(* Logix 5000 project; controller CIP_14485201 vendor 1 type 14 code 216 rev 38.11; software revision 38.01; part 9 of 12 *)
(* tags used below, declared in another part *)
   Bit : BOOL[128];   // BIT
   MOA_OFF : DINT[20];   // PANELVIEW MOA OFF
   MOA_ON : DINT[20];   // PANELVIEW MOA ON
   OpCode_Pin : DINT[5];   // OPCODE PIN ARRAY
   Panelview : INT[40];   // PANELVIEW CONTROL
   PID2 : PID;   // SUPPLY FLOW PID
   PID2_bumpless_transfer : BOOL;   // FORCE PID TO RESTART FROM PREVIOUS OUTPUT VALUE
   PID2_Man_Mode : BOOL;   // PID2 MANUAL MODE
   PID2_Manual_PB_Pressed : BOOL;   // PID2 MANUAL PUSHBUTTON PRESSED
   PID2_Output_Memory : REAL;   // SUPPLY FLOW PID OUTPUT MEMORY TO USE FOR BUMPLESS TRANSFER
   PID2_PV_Manual_PB : BOOL;   // PID2 MANUAL MODE SELECTED ON HMI
   PID2_Setpoint_Memory : REAL;   // SUPPLY FLOW PID SETPOINT MEMORY TO USE FOR BUMPLESS TRANSFER
   PID_Ons : DINT[6];   // PID ONE SHOT
   PID_Timer : TIMER[5];   // PID TIMERS
   PV_Output_Status : INT[20];   // PV OUTPUT STATUS:
   PV_Output_Status_IND : INT[20,16];   // PV OUTPUT STATUS IND:
   PV_Status_Bit : BOOL;   // SYSTEM BIT
   Recipe : RECIPE[41];   // RECIPES
   SP_Supply_Flow : REAL;   // CURRENT SUPPLY FLOW SETPOINT
   Supply_Mod_Valve_force_open : BOOL;   // FORCE SUPPLY MOD. VALVE TO 100% OPEN
   Utility_Button : DINT[5];   // PANELVIEW UTILITY BUTTONS
   Utility_Button_Ons : DINT[5];   // PANELVIEW UTILITY BUTTON ONE SHOTS
   Utility_Ons : DINT[5];   // PANELVIEW UTILITY ONE SHOTS
   Utility_Out : DINT[5];   // PANELVIEW UTILITY OUTPUT CONTROL
   Utility_Timer : TIMER[4];   // PANELVIEW UTILITY TIMERS
(* MainProgram, continued *)

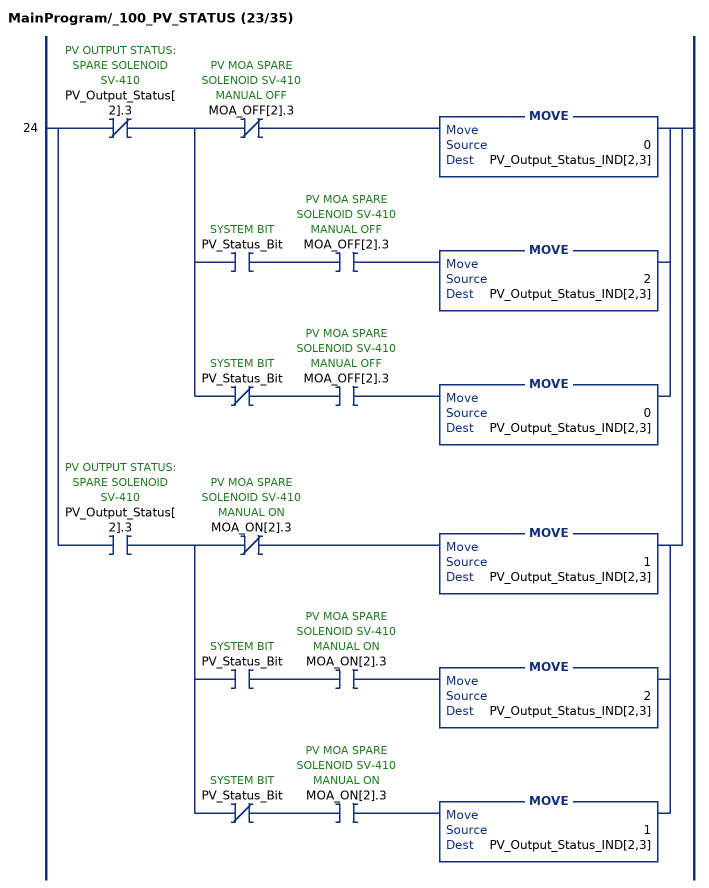
   [picture p140: MainProgram/_100_PV_STATUS rungs 24-24]
   24: [XIO(PV_Output_Status[2].3) [XIO(MOA_OFF[2].3) MOVE(0,PV_Output_Status_IND[2,3]) ,XIC(PV_Status_Bit) XIC(MOA_OFF[2].3) MOVE(2,PV_Output_Status_IND[2,3]) ,XIO(PV_Status_Bit) XIC(MOA_OFF[2].3) MOVE(0,PV_Output_Status_IND[2,3]) ] ,XIC(PV_Output_Status[2].3) [XIO(MOA_ON[2].3) MOVE(1,PV_Output_Status_IND[2,3]) ,XIC(PV_Status_Bit) XIC(MOA_ON[2].3) MOVE(2,PV_Output_Status_IND[2,3]) ,XIO(PV_Status_Bit) XIC(MOA_ON[2].3) MOVE(1,PV_Output_Status_IND[2,3]) ] ];
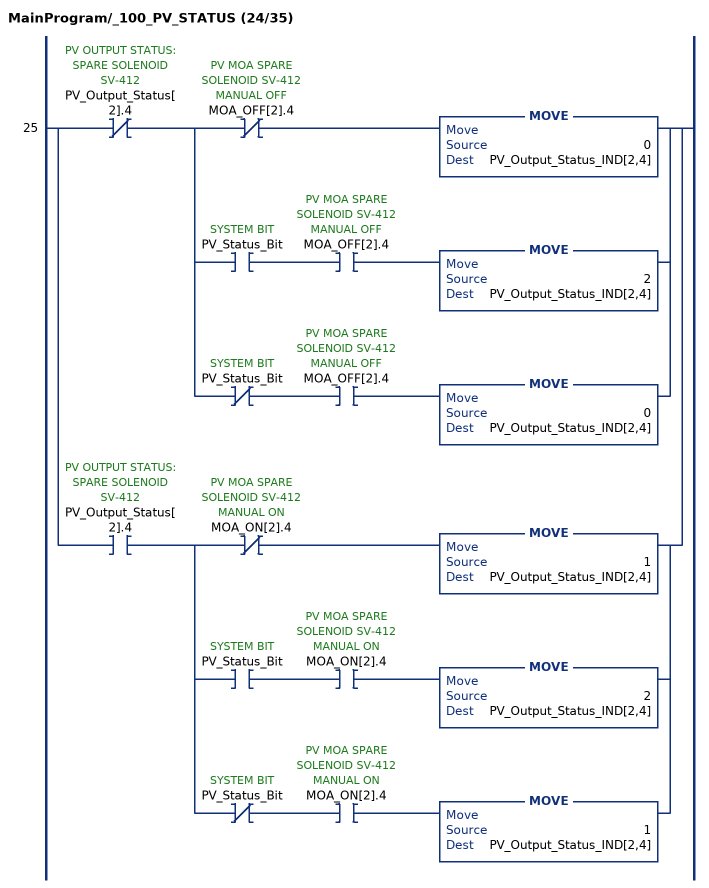
   25: [XIO(PV_Output_Status[2].4) [XIO(MOA_OFF[2].4) MOVE(0,PV_Output_Status_IND[2,4]) ,XIC(PV_Status_Bit) XIC(MOA_OFF[2].4) MOVE(2,PV_Output_Status_IND[2,4]) ,XIO(PV_Status_Bit) XIC(MOA_OFF[2].4) MOVE(0,PV_Output_Status_IND[2,4]) ] ,XIC(PV_Output_Status[2].4) [XIO(MOA_ON[2].4) MOVE(1,PV_Output_Status_IND[2,4]) ,XIC(PV_Status_Bit) XIC(MOA_ON[2].4) MOVE(2,PV_Output_Status_IND[2,4]) ,XIO(PV_Status_Bit) XIC(MOA_ON[2].4) MOVE(1,PV_Output_Status_IND[2,4]) ] ];
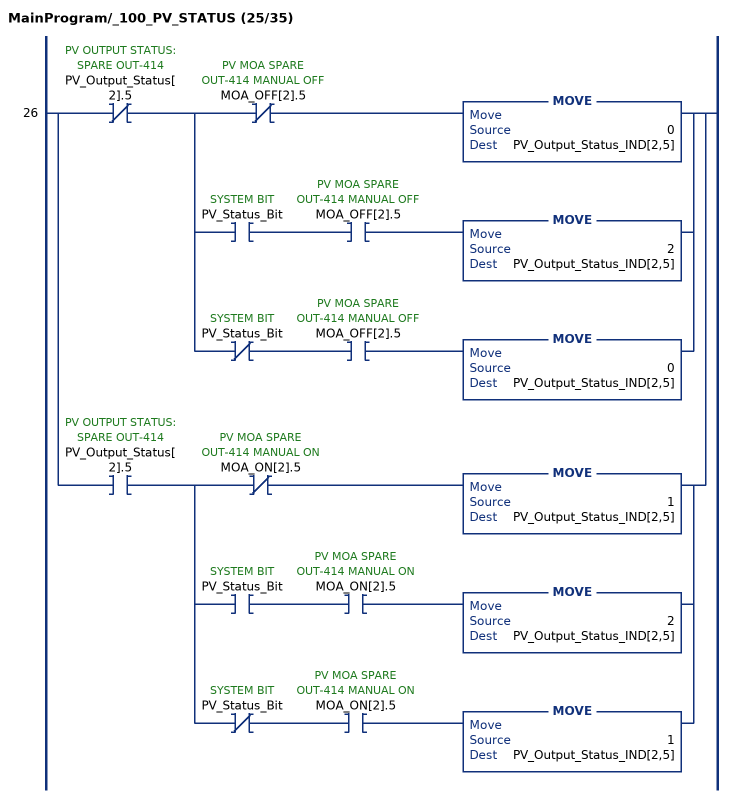
   26: [XIO(PV_Output_Status[2].5) [XIO(MOA_OFF[2].5) MOVE(0,PV_Output_Status_IND[2,5]) ,XIC(PV_Status_Bit) XIC(MOA_OFF[2].5) MOVE(2,PV_Output_Status_IND[2,5]) ,XIO(PV_Status_Bit) XIC(MOA_OFF[2].5) MOVE(0,PV_Output_Status_IND[2,5]) ] ,XIC(PV_Output_Status[2].5) [XIO(MOA_ON[2].5) MOVE(1,PV_Output_Status_IND[2,5]) ,XIC(PV_Status_Bit) XIC(MOA_ON[2].5) MOVE(2,PV_Output_Status_IND[2,5]) ,XIO(PV_Status_Bit) XIC(MOA_ON[2].5) MOVE(1,PV_Output_Status_IND[2,5]) ] ];
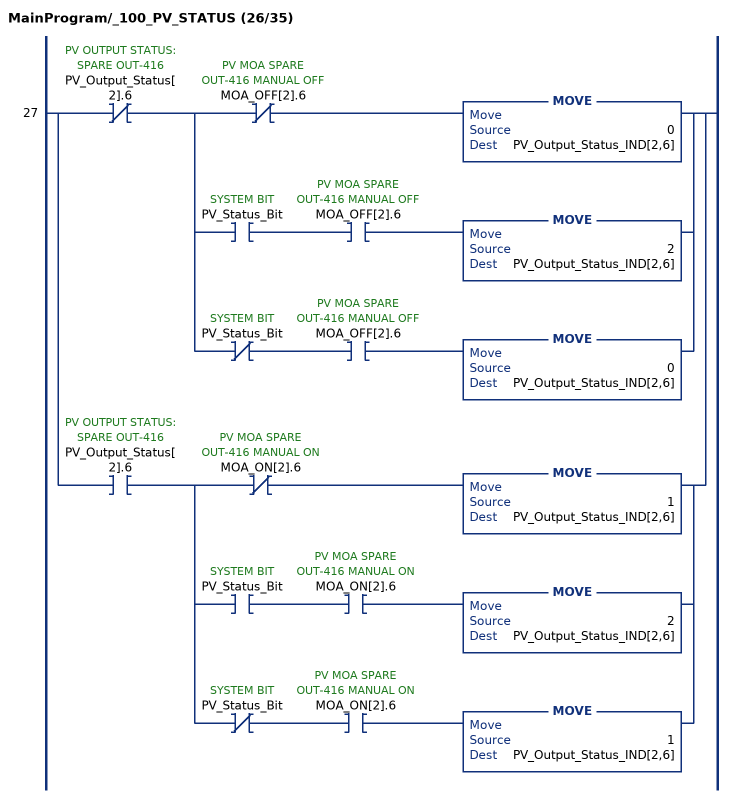
   27: [XIO(PV_Output_Status[2].6) [XIO(MOA_OFF[2].6) MOVE(0,PV_Output_Status_IND[2,6]) ,XIC(PV_Status_Bit) XIC(MOA_OFF[2].6) MOVE(2,PV_Output_Status_IND[2,6]) ,XIO(PV_Status_Bit) XIC(MOA_OFF[2].6) MOVE(0,PV_Output_Status_IND[2,6]) ] ,XIC(PV_Output_Status[2].6) [XIO(MOA_ON[2].6) MOVE(1,PV_Output_Status_IND[2,6]) ,XIC(PV_Status_Bit) XIC(MOA_ON[2].6) MOVE(2,PV_Output_Status_IND[2,6]) ,XIO(PV_Status_Bit) XIC(MOA_ON[2].6) MOVE(1,PV_Output_Status_IND[2,6]) ] ];
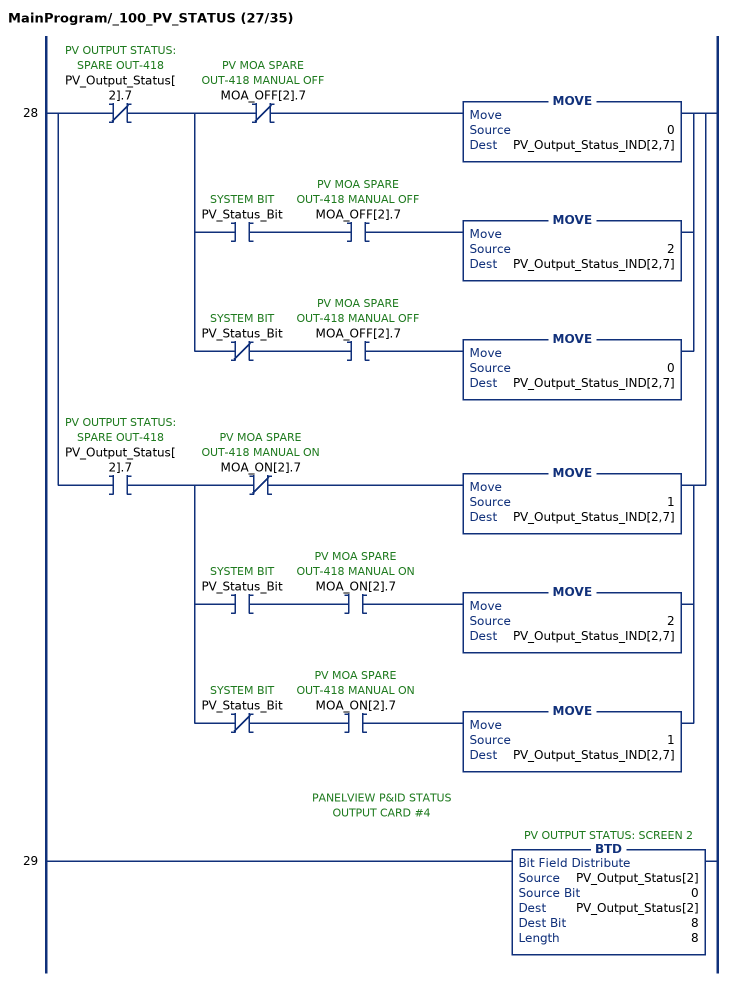
   28: [XIO(PV_Output_Status[2].7) [XIO(MOA_OFF[2].7) MOVE(0,PV_Output_Status_IND[2,7]) ,XIC(PV_Status_Bit) XIC(MOA_OFF[2].7) MOVE(2,PV_Output_Status_IND[2,7]) ,XIO(PV_Status_Bit) XIC(MOA_OFF[2].7) MOVE(0,PV_Output_Status_IND[2,7]) ] ,XIC(PV_Output_Status[2].7) [XIO(MOA_ON[2].7) MOVE(1,PV_Output_Status_IND[2,7]) ,XIC(PV_Status_Bit) XIC(MOA_ON[2].7) MOVE(2,PV_Output_Status_IND[2,7]) ,XIO(PV_Status_Bit) XIC(MOA_ON[2].7) MOVE(1,PV_Output_Status_IND[2,7]) ] ];
   // PANELVIEW P&ID STATUS
   // OUTPUT CARD #4
   29: BTD(PV_Output_Status[2],0,PV_Output_Status[2],8,8);
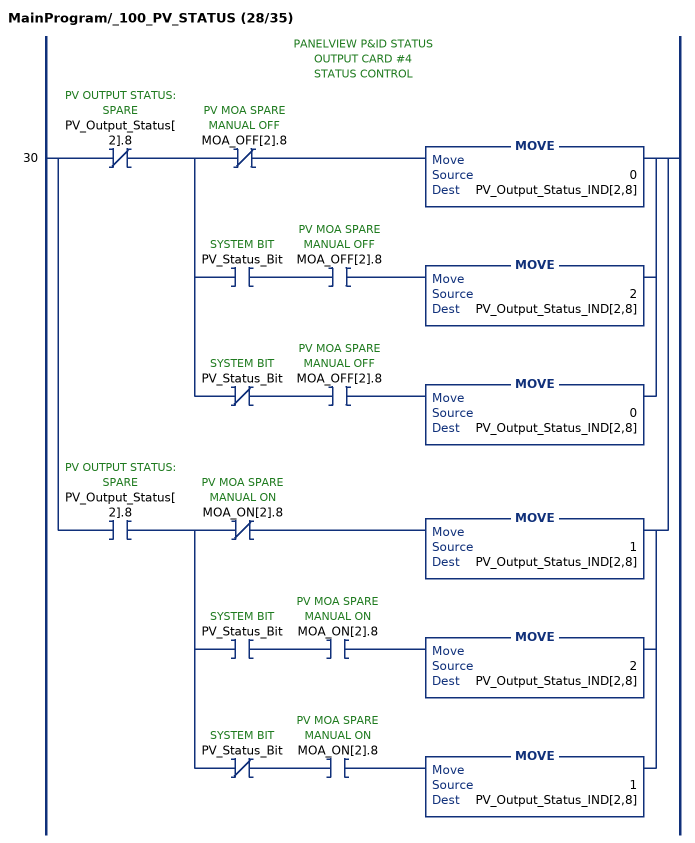
   // PANELVIEW P&ID STATUS
   // OUTPUT CARD #4
   // STATUS CONTROL
   30: [XIO(PV_Output_Status[2].8) [XIO(MOA_OFF[2].8) MOVE(0,PV_Output_Status_IND[2,8]) ,XIC(PV_Status_Bit) XIC(MOA_OFF[2].8) MOVE(2,PV_Output_Status_IND[2,8]) ,XIO(PV_Status_Bit) XIC(MOA_OFF[2].8) MOVE(0,PV_Output_Status_IND[2,8]) ] ,XIC(PV_Output_Status[2].8) [XIO(MOA_ON[2].8) MOVE(1,PV_Output_Status_IND[2,8]) ,XIC(PV_Status_Bit) XIC(MOA_ON[2].8) MOVE(2,PV_Output_Status_IND[2,8]) ,XIO(PV_Status_Bit) XIC(MOA_ON[2].8) MOVE(1,PV_Output_Status_IND[2,8]) ] ];
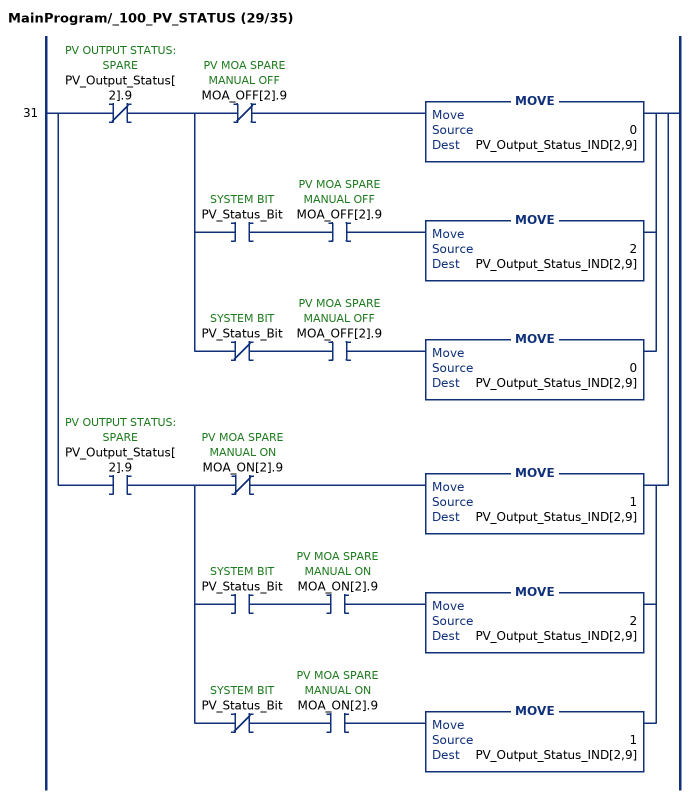
   31: [XIO(PV_Output_Status[2].9) [XIO(MOA_OFF[2].9) MOVE(0,PV_Output_Status_IND[2,9]) ,XIC(PV_Status_Bit) XIC(MOA_OFF[2].9) MOVE(2,PV_Output_Status_IND[2,9]) ,XIO(PV_Status_Bit) XIC(MOA_OFF[2].9) MOVE(0,PV_Output_Status_IND[2,9]) ] ,XIC(PV_Output_Status[2].9) [XIO(MOA_ON[2].9) MOVE(1,PV_Output_Status_IND[2,9]) ,XIC(PV_Status_Bit) XIC(MOA_ON[2].9) MOVE(2,PV_Output_Status_IND[2,9]) ,XIO(PV_Status_Bit) XIC(MOA_ON[2].9) MOVE(1,PV_Output_Status_IND[2,9]) ] ];
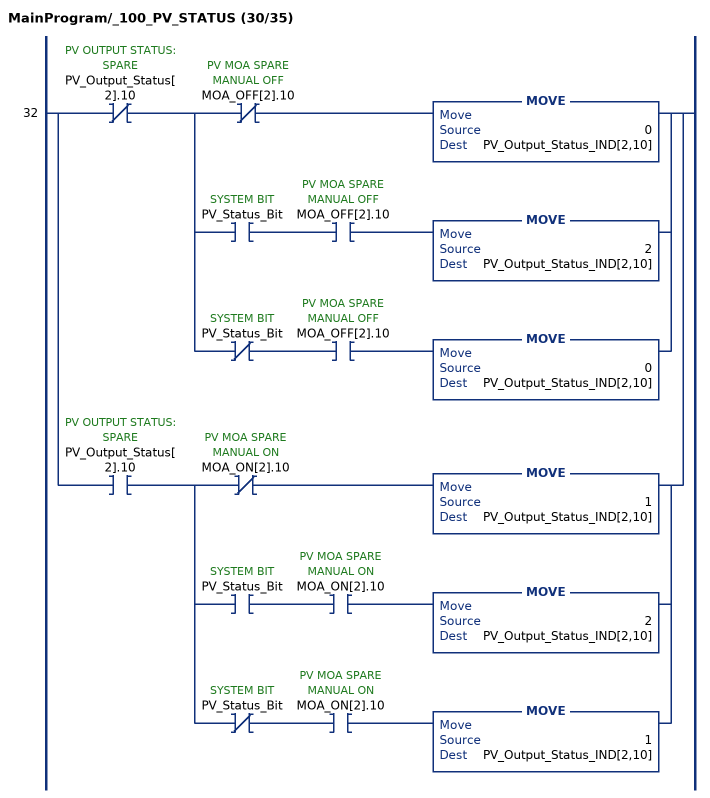
   32: [XIO(PV_Output_Status[2].10) [XIO(MOA_OFF[2].10) MOVE(0,PV_Output_Status_IND[2,10]) ,XIC(PV_Status_Bit) XIC(MOA_OFF[2].10) MOVE(2,PV_Output_Status_IND[2,10]) ,XIO(PV_Status_Bit) XIC(MOA_OFF[2].10) MOVE(0,PV_Output_Status_IND[2,10]) ] ,XIC(PV_Output_Status[2].10) [XIO(MOA_ON[2].10) MOVE(1,PV_Output_Status_IND[2,10]) ,XIC(PV_Status_Bit) XIC(MOA_ON[2].10) MOVE(2,PV_Output_Status_IND[2,10]) ,XIO(PV_Status_Bit) XIC(MOA_ON[2].10) MOVE(1,PV_Output_Status_IND[2,10]) ] ];
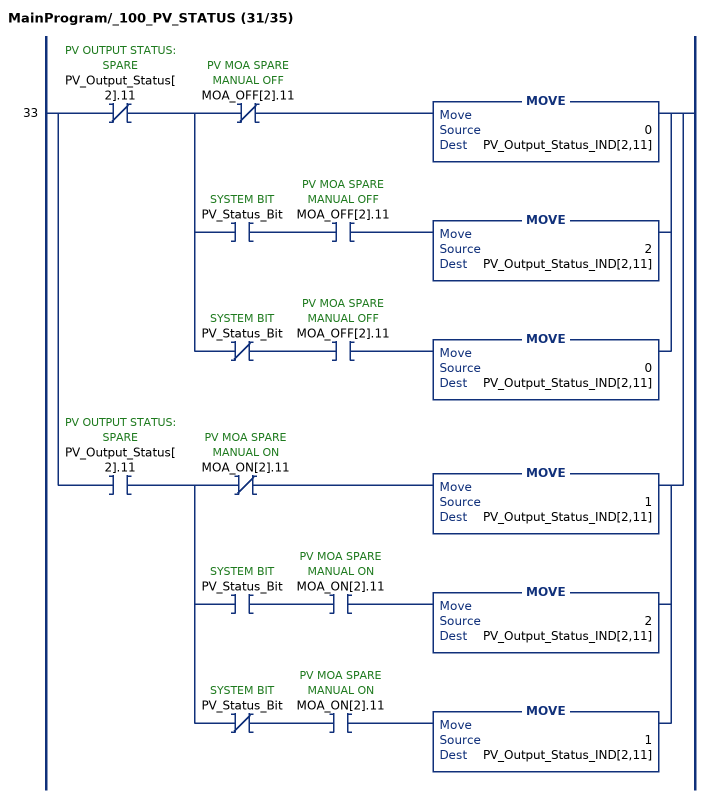
   33: [XIO(PV_Output_Status[2].11) [XIO(MOA_OFF[2].11) MOVE(0,PV_Output_Status_IND[2,11]) ,XIC(PV_Status_Bit) XIC(MOA_OFF[2].11) MOVE(2,PV_Output_Status_IND[2,11]) ,XIO(PV_Status_Bit) XIC(MOA_OFF[2].11) MOVE(0,PV_Output_Status_IND[2,11]) ] ,XIC(PV_Output_Status[2].11) [XIO(MOA_ON[2].11) MOVE(1,PV_Output_Status_IND[2,11]) ,XIC(PV_Status_Bit) XIC(MOA_ON[2].11) MOVE(2,PV_Output_Status_IND[2,11]) ,XIO(PV_Status_Bit) XIC(MOA_ON[2].11) MOVE(1,PV_Output_Status_IND[2,11]) ] ];
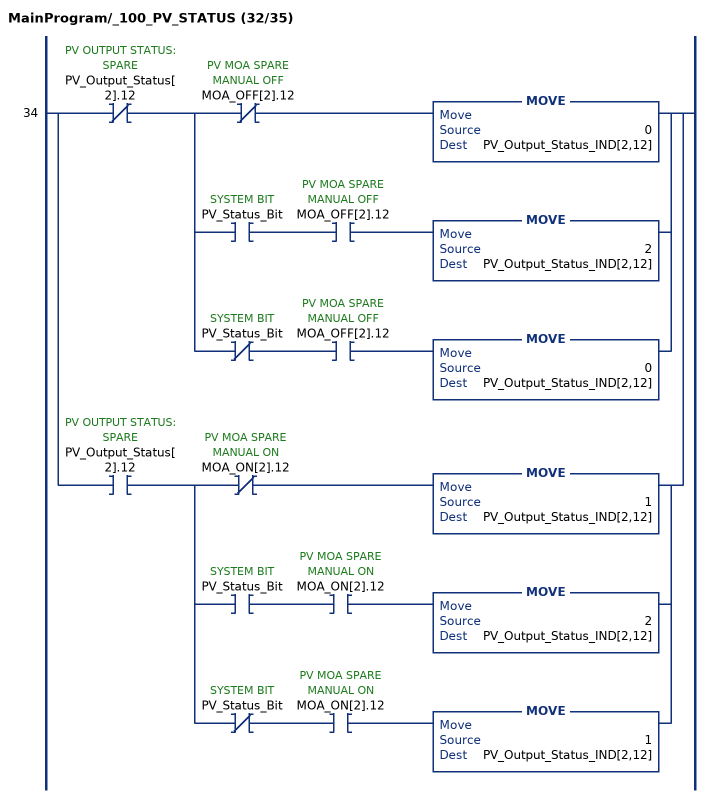
   34: [XIO(PV_Output_Status[2].12) [XIO(MOA_OFF[2].12) MOVE(0,PV_Output_Status_IND[2,12]) ,XIC(PV_Status_Bit) XIC(MOA_OFF[2].12) MOVE(2,PV_Output_Status_IND[2,12]) ,XIO(PV_Status_Bit) XIC(MOA_OFF[2].12) MOVE(0,PV_Output_Status_IND[2,12]) ] ,XIC(PV_Output_Status[2].12) [XIO(MOA_ON[2].12) MOVE(1,PV_Output_Status_IND[2,12]) ,XIC(PV_Status_Bit) XIC(MOA_ON[2].12) MOVE(2,PV_Output_Status_IND[2,12]) ,XIO(PV_Status_Bit) XIC(MOA_ON[2].12) MOVE(1,PV_Output_Status_IND[2,12]) ] ];
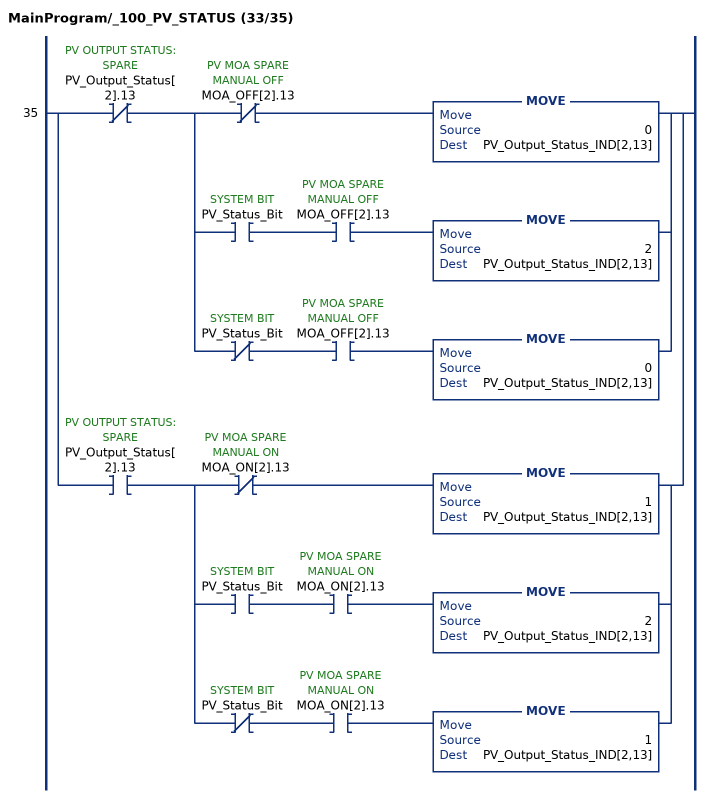
   35: [XIO(PV_Output_Status[2].13) [XIO(MOA_OFF[2].13) MOVE(0,PV_Output_Status_IND[2,13]) ,XIC(PV_Status_Bit) XIC(MOA_OFF[2].13) MOVE(2,PV_Output_Status_IND[2,13]) ,XIO(PV_Status_Bit) XIC(MOA_OFF[2].13) MOVE(0,PV_Output_Status_IND[2,13]) ] ,XIC(PV_Output_Status[2].13) [XIO(MOA_ON[2].13) MOVE(1,PV_Output_Status_IND[2,13]) ,XIC(PV_Status_Bit) XIC(MOA_ON[2].13) MOVE(2,PV_Output_Status_IND[2,13]) ,XIO(PV_Status_Bit) XIC(MOA_ON[2].13) MOVE(1,PV_Output_Status_IND[2,13]) ] ];
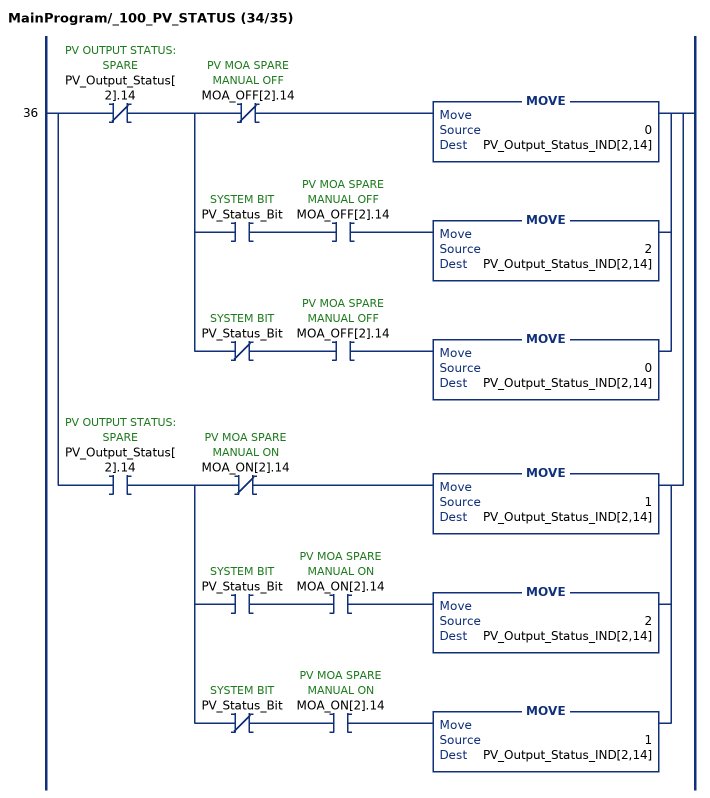
   36: [XIO(PV_Output_Status[2].14) [XIO(MOA_OFF[2].14) MOVE(0,PV_Output_Status_IND[2,14]) ,XIC(PV_Status_Bit) XIC(MOA_OFF[2].14) MOVE(2,PV_Output_Status_IND[2,14]) ,XIO(PV_Status_Bit) XIC(MOA_OFF[2].14) MOVE(0,PV_Output_Status_IND[2,14]) ] ,XIC(PV_Output_Status[2].14) [XIO(MOA_ON[2].14) MOVE(1,PV_Output_Status_IND[2,14]) ,XIC(PV_Status_Bit) XIC(MOA_ON[2].14) MOVE(2,PV_Output_Status_IND[2,14]) ,XIO(PV_Status_Bit) XIC(MOA_ON[2].14) MOVE(1,PV_Output_Status_IND[2,14]) ] ];
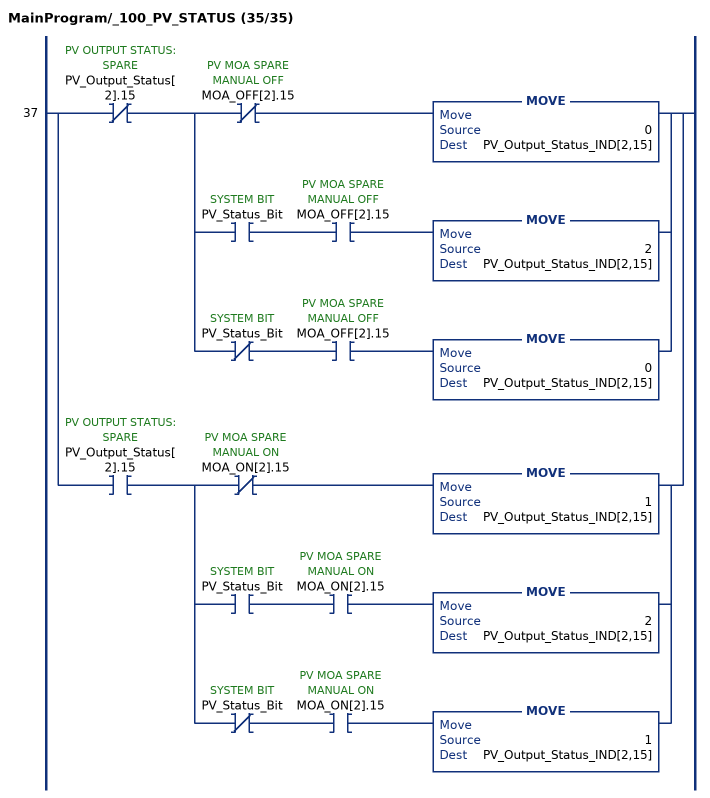
   37: [XIO(PV_Output_Status[2].15) [XIO(MOA_OFF[2].15) MOVE(0,PV_Output_Status_IND[2,15]) ,XIC(PV_Status_Bit) XIC(MOA_OFF[2].15) MOVE(2,PV_Output_Status_IND[2,15]) ,XIO(PV_Status_Bit) XIC(MOA_OFF[2].15) MOVE(0,PV_Output_Status_IND[2,15]) ] ,XIC(PV_Output_Status[2].15) [XIO(MOA_ON[2].15) MOVE(1,PV_Output_Status_IND[2,15]) ,XIC(PV_Status_Bit) XIC(MOA_ON[2].15) MOVE(2,PV_Output_Status_IND[2,15]) ,XIO(PV_Status_Bit) XIC(MOA_ON[2].15) MOVE(1,PV_Output_Status_IND[2,15]) ] ];
END_ROUTINE

ROUTINE _20_UTILITY   (* ladder *)
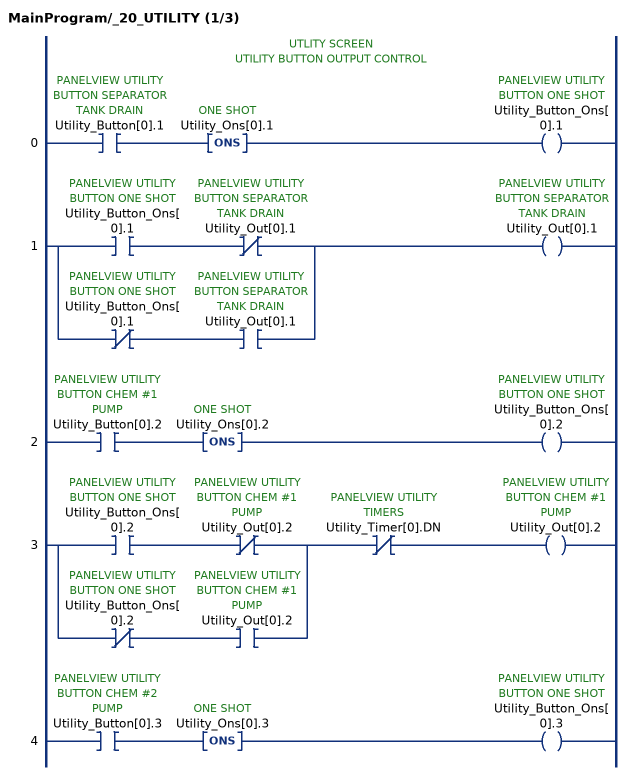
   // UTLITY SCREEN
   // UTILITY BUTTON OUTPUT CONTROL
   0: XIC(Utility_Button[0].1)ONS(Utility_Ons[0].1)OTE(Utility_Button_Ons[0].1);
   1: [XIC(Utility_Button_Ons[0].1) XIO(Utility_Out[0].1) ,XIO(Utility_Button_Ons[0].1) XIC(Utility_Out[0].1) ]OTE(Utility_Out[0].1);
   2: XIC(Utility_Button[0].2)ONS(Utility_Ons[0].2)OTE(Utility_Button_Ons[0].2);
   3: [XIC(Utility_Button_Ons[0].2) XIO(Utility_Out[0].2) ,XIO(Utility_Button_Ons[0].2) XIC(Utility_Out[0].2) ]XIO(Utility_Timer[0].DN)OTE(Utility_Out[0].2);
   4: XIC(Utility_Button[0].3)ONS(Utility_Ons[0].3)OTE(Utility_Button_Ons[0].3);
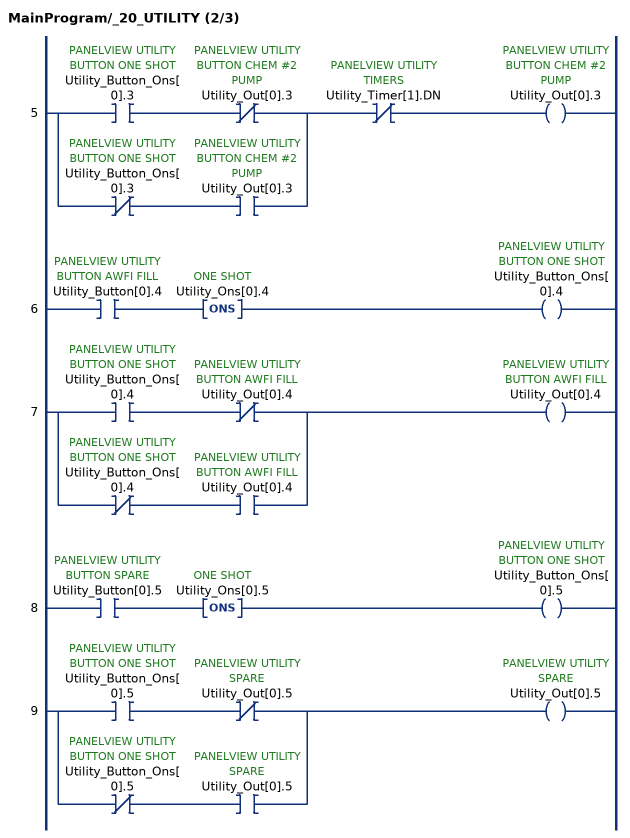
   5: [XIC(Utility_Button_Ons[0].3) XIO(Utility_Out[0].3) ,XIO(Utility_Button_Ons[0].3) XIC(Utility_Out[0].3) ]XIO(Utility_Timer[1].DN)OTE(Utility_Out[0].3);
   6: XIC(Utility_Button[0].4)ONS(Utility_Ons[0].4)OTE(Utility_Button_Ons[0].4);
   7: [XIC(Utility_Button_Ons[0].4) XIO(Utility_Out[0].4) ,XIO(Utility_Button_Ons[0].4) XIC(Utility_Out[0].4) ]OTE(Utility_Out[0].4);
   8: XIC(Utility_Button[0].5)ONS(Utility_Ons[0].5)OTE(Utility_Button_Ons[0].5);
   9: [XIC(Utility_Button_Ons[0].5) XIO(Utility_Out[0].5) ,XIO(Utility_Button_Ons[0].5) XIC(Utility_Out[0].5) ]OTE(Utility_Out[0].5);
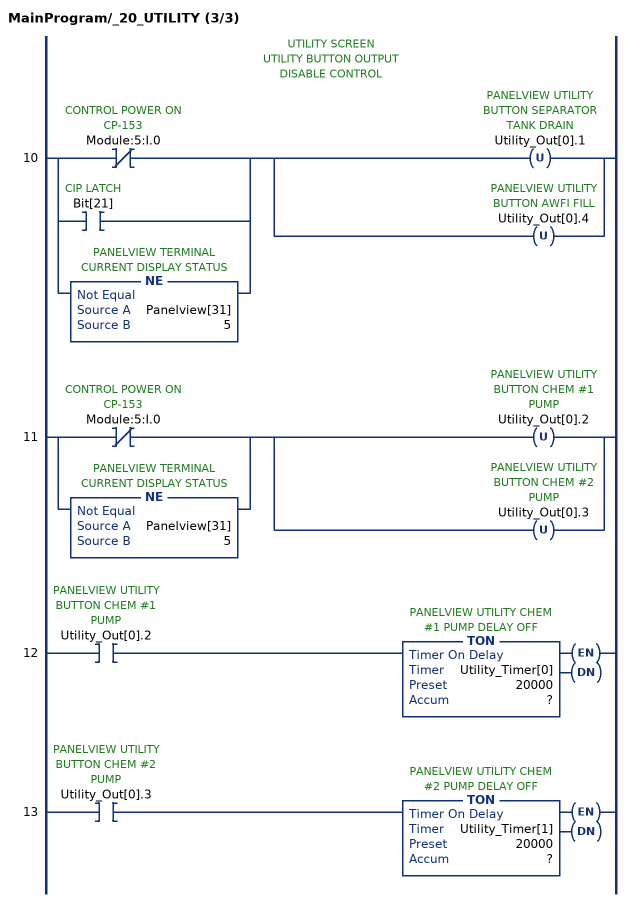
   // UTILITY SCREEN
   // UTILITY BUTTON OUTPUT
   // DISABLE CONTROL
   10: [XIO(Module:5:I.0) ,XIC(Bit[21]) ,NE(Panelview[31],5) ][OTU(Utility_Out[0].1) ,OTU(Utility_Out[0].4) ];
   11: [XIO(Module:5:I.0) ,NE(Panelview[31],5) ][OTU(Utility_Out[0].2) ,OTU(Utility_Out[0].3) ];
   12: XIC(Utility_Out[0].2)TON(Utility_Timer[0],?,?);
   13: XIC(Utility_Out[0].3)TON(Utility_Timer[1],?,?);
END_ROUTINE

ROUTINE _25_PID_SUPPLY_FLOW   (* ladder *)
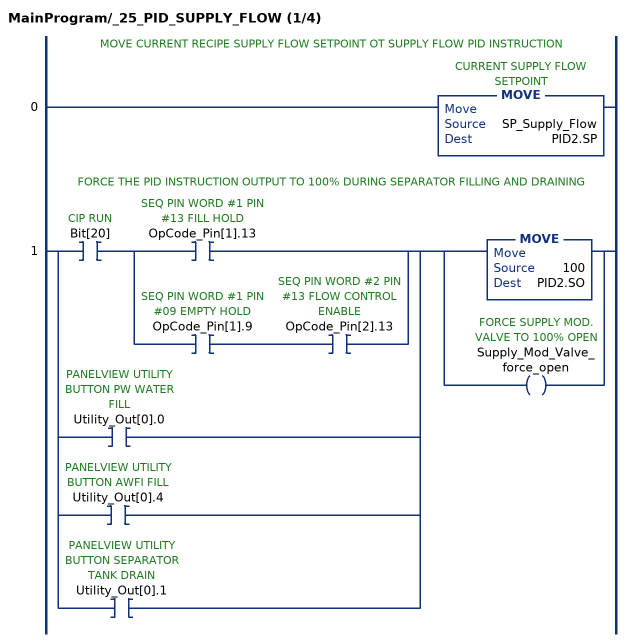
   // MOVE CURRENT RECIPE SUPPLY FLOW SETPOINT OT SUPPLY FLOW PID INSTRUCTION
   0: MOVE(SP_Supply_Flow,PID2.SP);
   // FORCE THE PID INSTRUCTION OUTPUT TO 100% DURING SEPARATOR FILLING AND DRAINING
   1: [XIC(Bit[20]) [XIC(OpCode_Pin[1].13) ,XIC(OpCode_Pin[1].9) XIC(OpCode_Pin[2].13) ] ,XIC(Utility_Out[0].0) ,XIC(Utility_Out[0].4) ,XIC(Utility_Out[0].1) ][MOVE(100,PID2.SO) ,OTE(Supply_Mod_Valve_force_open) ];
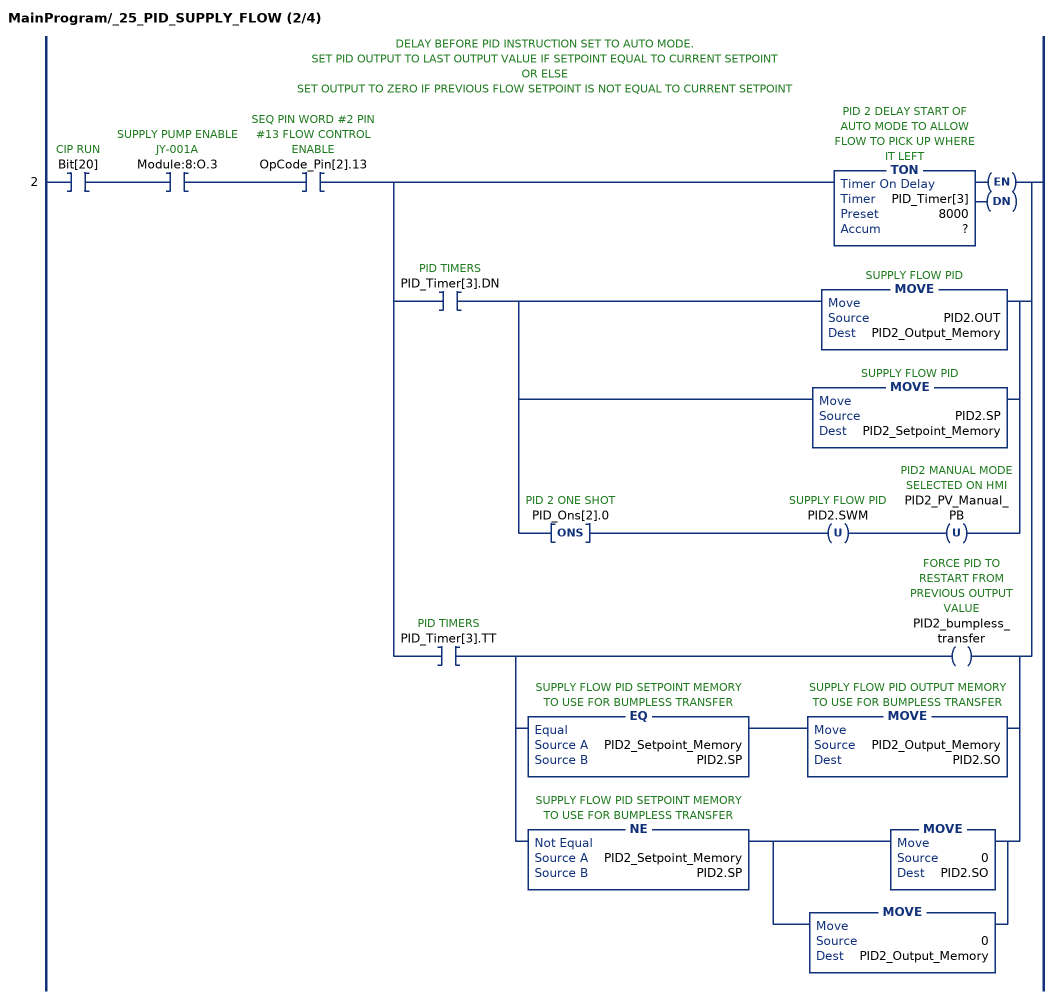
   // DELAY BEFORE PID INSTRUCTION SET TO AUTO MODE.
   // SET PID OUTPUT TO LAST OUTPUT VALUE IF SETPOINT EQUAL TO CURRENT SETPOINT
   // OR ELSE
   // SET OUTPUT TO ZERO IF PREVIOUS FLOW SETPOINT IS NOT EQUAL TO CURRENT SETPOINT
   2: XIC(Bit[20])XIC(Module:8:O.3)XIC(OpCode_Pin[2].13)[TON(PID_Timer[3],?,?) ,XIC(PID_Timer[3].DN) [MOVE(PID2.OUT,PID2_Output_Memory) ,MOVE(PID2.SP,PID2_Setpoint_Memory) ,ONS(PID_Ons[2].0) OTU(PID2.SWM) OTU(PID2_PV_Manual_PB) ] ,XIC(PID_Timer[3].TT) [OTE(PID2_bumpless_transfer) ,EQ(PID2_Setpoint_Memory,PID2.SP) MOVE(PID2_Output_Memory,PID2.SO) ,NE(PID2_Setpoint_Memory,PID2.SP) [MOVE(0,PID2.SO) ,MOVE(0,PID2_Output_Memory) ] ] ];
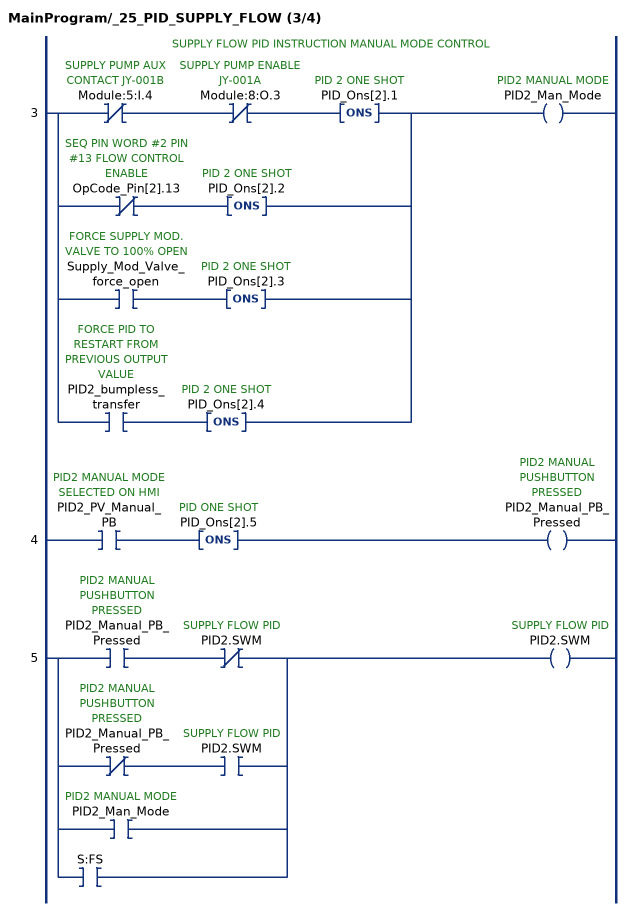
   // SUPPLY FLOW PID INSTRUCTION MANUAL MODE CONTROL
   3: [XIO(Module:5:I.4) XIO(Module:8:O.3) ONS(PID_Ons[2].1) ,XIO(OpCode_Pin[2].13) ONS(PID_Ons[2].2) ,XIC(Supply_Mod_Valve_force_open) ONS(PID_Ons[2].3) ,XIC(PID2_bumpless_transfer) ONS(PID_Ons[2].4) ]OTE(PID2_Man_Mode);
   4: XIC(PID2_PV_Manual_PB)ONS(PID_Ons[2].5)OTE(PID2_Manual_PB_Pressed);
   5: [XIC(PID2_Manual_PB_Pressed) XIO(PID2.SWM) ,XIO(PID2_Manual_PB_Pressed) XIC(PID2.SWM) ,XIC(PID2_Man_Mode) ,XIC(S:FS) ]OTE(PID2.SWM);
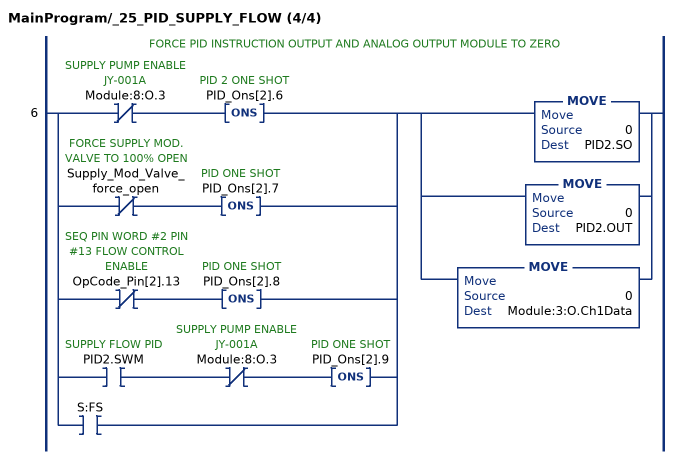
   // FORCE PID INSTRUCTION OUTPUT AND ANALOG OUTPUT MODULE TO ZERO
   6: [XIO(Module:8:O.3) ONS(PID_Ons[2].6) ,XIO(Supply_Mod_Valve_force_open) ONS(PID_Ons[2].7) ,XIO(OpCode_Pin[2].13) ONS(PID_Ons[2].8) ,XIC(PID2.SWM) XIO(Module:8:O.3) ONS(PID_Ons[2].9) ,XIC(S:FS) ][MOVE(0,PID2.SO) ,MOVE(0,PID2.OUT) ,MOVE(0,Module:3:O.Ch1Data) ];
END_ROUTINE
